Fanuc KAREL source: kb00189.compact.KL

PROGRAM KB00189
%STACKSIZE=65535
%PRIORITY=65535
%NOLOCKGROUP
VAR
P1 : STRING[80]
P2 : INTEGER
P3 : INTEGER
RESULT : STRING[80]
BEGIN
P1='A'
P2=1
P3=1
RESULT=SUB_STR(P1,P2,P3)
END KB00189
